(* IEC 61131-3 sources: kns-port-domestic/tools/port_metrics_tests/fixtures/adapted/src/DUTs, 2 files *)

(* ---- E_PumpMode.dut.st ---- *)
{attribute 'qualified_only'}
{attribute 'strict'}
TYPE E_PumpMode :
(
    Auto := 1,
    Manual := 2
); // PORT: [types] перечисление без базового типа (F34)
END_TYPE

(* ---- ST_PumpCfg.dut.st ---- *)
TYPE ST_PumpCfg :
STRUCT
    rSpeedMax_Hz : REAL := 50.0; // предел частоты, Гц
    tStartDelay : TIME := T#5S;
END_STRUCT
END_TYPE
